PROGRAM MAIN
VAR
	i: INT;
	ton_TwinSAFE_ACK_reset: TON;
	BlinkLED: ton;

	Pulse_On_TON: TON;
	Pulse_Off_TON: TON;
	bPulse	:	BOOL	;
	
	t_BlinkTime : TIME	;
	
	n_SafeSate	:	INT	;
END_VAR

i:=i+1;


ton_TwinSAFE_ACK_reset(IN:=GVL_Safety.stTwinSAFE_OUT.ErrACK, PT:=T#10S);
IF ton_TwinSAFE_ACK_reset.Q THEN;
	GVL_Safety.stTwinSAFE_OUT.ErrACK:=FALSE;
END_IF
GVL_Safety.stTwinSAFE_OUT.DoorMonitor:=GVL_Safety.DoorMonitorFromPLC;

//Battery Relay CMD
IF GVL_Safety.stTwinSAFE_OUT.BatRelay_CMD THEN
	GVL_Safety.stTwinSAFE_OUT.BatRelay_Manual_Off:=FALSE;
	GVL_Safety.stTwinSAFE_OUT.BatRelay_Manual_On:=TRUE;
ELSE
	GVL_Safety.stTwinSAFE_OUT.BatRelay_Manual_Off:=TRUE;
	GVL_Safety.stTwinSAFE_OUT.BatRelay_Manual_On:=FALSE;
END_IF

//Battery BMS Relay CMD
IF GVL_Safety.stTwinSAFE_OUT.BatBMS_Cmd THEN
	GVL_Safety.stTwinSAFE_OUT.RB_BatBMS_Manual_Off:=FALSE;
	GVL_Safety.stTwinSAFE_OUT.RB_BatBMS_Manual_On:=TRUE;
ELSE
	GVL_Safety.stTwinSAFE_OUT.RB_BatBMS_Manual_Off:=TRUE;
	GVL_Safety.stTwinSAFE_OUT.RB_BatBMS_Manual_On:=FALSE;

END_IF

act_LED_Control();
act_LogicMap();

ACTION act_LED_Control:
//Red 
IF GVL_Safety.stTwinSAFE_IN.EStop_Ok AND GVL_Safety.stTwinSAFE_IN.EStop_Status THEN
	//Red Off
	GVL_IO.RedLED:= FALSE;
ELSIF GVL_Safety.stTwinSAFE_IN.EStop_Ok=FALSE AND GVL_Safety.stTwinSAFE_IN.EStop_Status  THEN
	//Red Blink 
	GVL_IO.RedLED:=bPulse;
ELSIF GVL_Safety.stTwinSAFE_IN.EStop_Ok=FALSE AND GVL_Safety.stTwinSAFE_IN.EStop_Status=FALSE THEN
	//Red On
	GVL_IO.RedLED:= TRUE;
END_IF

//Blue
IF (GVL_Safety.stTwinSAFE_OUT.DoorMonitor AND GVL_Safety.stTwinSAFE_IN.Speps.step1) 
OR (GVL_Safety.stTwinSAFE_OUT.DoorMonitor=FALSE AND GVL_Safety.stTwinSAFE_IN.Speps.stepRnD) THEN
	//Blue Blink
	GVL_IO.BlueLED:=bPulse;
ELSIF GVL_Safety.stTwinSAFE_OUT.DoorMonitor AND GVL_Safety.stTwinSAFE_OUT.SolenoedMonitor=FALSE AND NOT GVL_Safety.stTwinSAFE_IN.Speps.stepRnD THEN
	//Blue Off
	GVL_IO.BlueLED:=FALSE;
ELSIF GVL_Safety.stTwinSAFE_OUT.DoorMonitor=FALSE OR (GVL_Safety.stTwinSAFE_IN.Speps.stepRnD AND GVL_Safety.stTwinSAFE_OUT.DoorMonitor) THEN
	//Blue On
	GVL_IO.BlueLED:=TRUE;
END_IF

//Green
IF (GVL_Safety.stTwinSAFE_IN.Speps.step1 AND GVL_Safety.stTwinSAFE_IN.EStop_Ok AND GVL_Safety.stTwinSAFE_OUT.DoorMonitor=TRUE) OR GVL_Safety.stTwinSAFE_IN.TransitionStep THEN
	//Green Blink
	GVL_IO.GreenLED:=bPulse;
ELSIF GVL_Safety.stTwinSAFE_IN.Safety_Armed OR (GVL_Safety.stTwinSAFE_IN.Speps.stepRnD) OR GVL_Safety.stTwinSAFE_IN.Speps.step2 THEN
	//Green On
	GVL_IO.GreenLED:=TRUE;
ELSIF GVL_Safety.stTwinSAFE_IN.Speps.step4 OR GVL_Safety.stTwinSAFE_IN.Speps.step5 
OR GVL_Safety.stTwinSAFE_IN.Speps.step6 OR GVL_Safety.stTwinSAFE_OUT.DoorMonitor=FALSE THEN
	//Green Off
	GVL_IO.GreenLED:=FALSE;
END_IF

IF GVL_Safety.stTwinSAFE_IN.Speps.step2 OR GVL_Safety.stTwinSAFE_IN.TransitionStep THEN
	t_BlinkTime:=T#0.5S;
ELSE
	t_BlinkTime:=T#1.5S;
END_IF

Pulse_On_TON(IN:=NOT bPulse , PT:=t_BlinkTime , Q=> , ET=> );
Pulse_Off_TON(IN:=bPulse , PT:=t_BlinkTime , Q=> , ET=> );
IF Pulse_On_TON.Q AND NOT bPulse THEN bPulse:=TRUE; END_IF;
IF Pulse_Off_TON.Q AND bPulse THEN bPulse:=FALSE; END_IF;


GVL_Safety.stTwinSAFE_IN.HV_Healthy_Invert:=NOT GVL_Safety.stTwinSAFE_IN.HV_Healthy;
GVL_Safety.stTwinSAFE_IN.LV_Healthy_Invert:=NOT GVL_Safety.stTwinSAFE_IN.LV_Healthy;
END_ACTION

ACTION act_LogicMap:
(*
_________________________________________________________________________________________________________________________________________________________________
Function				|	Bit 1 (RnD Mode) GVL_Safety.stTwinSAFE_OUT.Set_RnD_Mode		|	Bit 2 (RnD Mode 2)		GVL_Safety.stTwinSAFE_OUT.Set_RnD_Mode2	|
________________________|_______________________________|_______________________________|
From Safe to RnD		|	1							|	0							|
________________________|_______________________________|_______________________________|
From RnD to Armed		|	1							|	1							|
________________________|_______________________________|_______________________________|
From RnD to Safe		|	0							|	0							|
________________________|_______________________________|_______________________________|
From Armed to RnD		|	0							|	1							|
________________________|_______________________________|_______________________________|

*)
;

GVL_Safety.stTwinSAFE_OUT.Set_RnD_Mode;
GVL_Safety.stTwinSAFE_OUT.Set_RnD_Mode2;

CASE n_SafeSate OF
	E_SafetyState.enum_RnD_2_Safe://From RnD to Safe	
		GVL_Safety.stTwinSAFE_OUT.Set_RnD_Mode:=FALSE;
		GVL_Safety.stTwinSAFE_OUT.Set_RnD_Mode2:=FALSE;
	E_SafetyState.enum_Safe_2_RnD://From Safe to RnD
		GVL_Safety.stTwinSAFE_OUT.Set_RnD_Mode:=TRUE;
		GVL_Safety.stTwinSAFE_OUT.Set_RnD_Mode2:=FALSE;
	
	E_SafetyState.enum_RnD_2_Armed://From RnD to Armed
		GVL_Safety.stTwinSAFE_OUT.Set_RnD_Mode:=TRUE;
		GVL_Safety.stTwinSAFE_OUT.Set_RnD_Mode2:=TRUE;
	
	E_SafetyState.enum_Armed_2_RnD://From Armed to RnD
		GVL_Safety.stTwinSAFE_OUT.Set_RnD_Mode:=TRUE;
		GVL_Safety.stTwinSAFE_OUT.Set_RnD_Mode2:=FALSE;
END_CASE


(*IF GVL_Safety.stTwinSAFE_OUT.Bypass_C1C2 THEN
	
END_IF*)
END_ACTION

END_PROGRAM

(* stored: Version 1.1.0.1, ProductVersion 3.1.4026.19
   POU MAIN: Id {0726ba31-cfa3-4f4b-8cfa-b894f8445811}, SpecialFunc None
   Action act_LED_Control: Id {3c867c17-f4c4-4546-bd10-836abda837f5}
   Action act_LogicMap: Id {0f0c44db-ccbd-41ab-9cfc-1e821c520f71} *)
